SUBAPPLICATION Uebung_268_AX (* Race Condition mit E_SPLIT: zwei falsche und zwei richtige Varianten (Adapter) *)
  (* Standard: 61499-2; Description: Copyright (c) 2026 Meisterschulen am Ostbahnhof This program and the accompanying materials are made available under the terms of the Eclipse Public License 2.0 which is available at https://www.eclipse.org/legal/epl-2.0/ SPDX-License-Identifier: EPL-2.0 *)
  (* Version 1.0, 2026-11-11, Franz Höpfinger, Meisterschulen am Ostbahnhof, initial API and implementation and/or initial documentation *)
  PACKAGE Uebungen;
  IMPORT logiBUS::io::DI::logiBUS_DI::Input_I1;
  IMPORT logiBUS::io::DI::logiBUS_DI::Input_I2;
  IMPORT logiBUS::io::DI::logiBUS_DI::Input_I3;
  IMPORT logiBUS::io::DI::logiBUS_DI::Input_I4;
  IMPORT logiBUS::io::DI::logiBUS_DI_Events::BUTTON_SINGLE_CLICK;
  IMPORT logiBUS::io::DQ::logiBUS_DO::Output_Q1;
  IMPORT logiBUS::io::DQ::logiBUS_DO::Output_Q2;
  IMPORT logiBUS::io::DQ::logiBUS_DO::Output_Q3;
  IMPORT logiBUS::io::DQ::logiBUS_DO::Output_Q4;
  IMPORT logiBUS::io::DQ::logiBUS_DO::Output_Q5;
  IMPORT logiBUS::io::DQ::logiBUS_DO::Output_Q6;
  IMPORT logiBUS::io::DQ::logiBUS_DO::Output_Q7;
  IMPORT logiBUS::io::DQ::logiBUS_DO::Output_Q8;
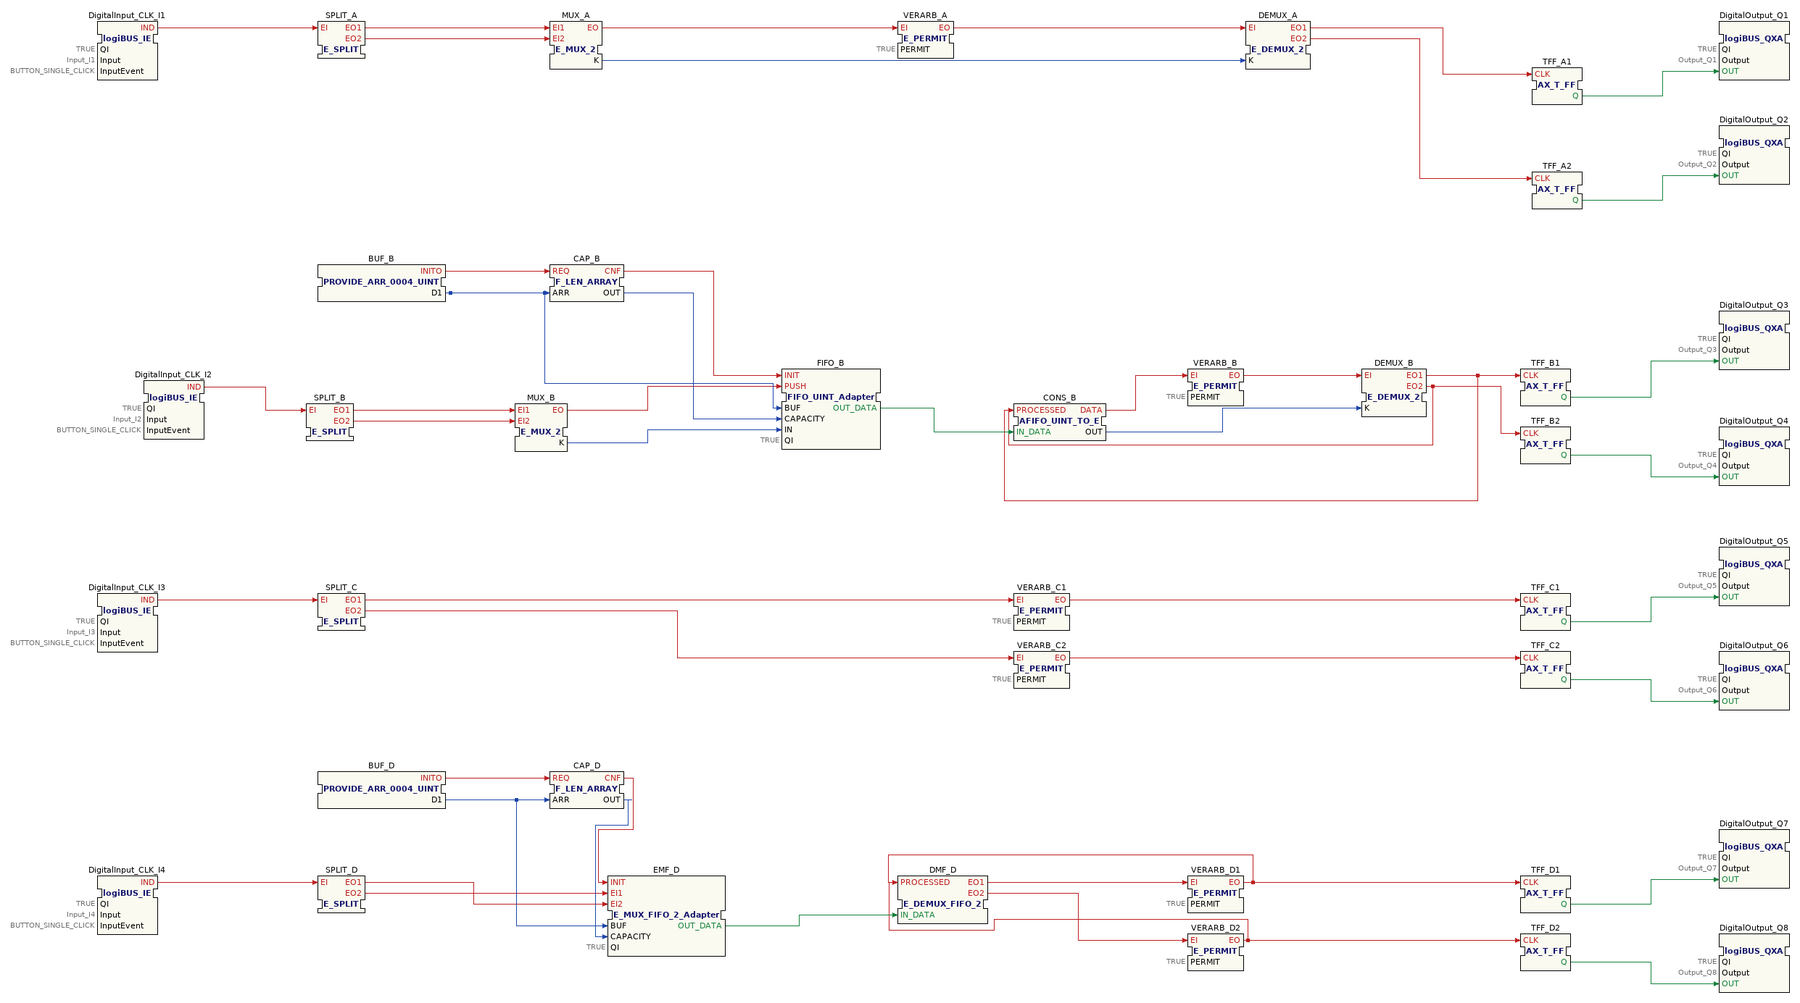
  FBS
    DigitalInput_CLK_I1 : logiBUS::io::DI::logiBUS_IE(QI := TRUE, Input := Input_I1, InputEvent := BUTTON_SINGLE_CLICK);
    SPLIT_A : iec61499::events::E_SPLIT;
    MUX_A : iec61499::events::E_MUX_2;
    VERARB_A : iec61499::events::E_PERMIT(PERMIT := TRUE);
    DEMUX_A : iec61499::events::E_DEMUX_2;
    TFF_A1 : adapter::events::unidirectional::AX_T_FF;
    DigitalOutput_Q1 : logiBUS::io::DQ::logiBUS_QXA(QI := TRUE, Output := Output_Q1);
    TFF_A2 : adapter::events::unidirectional::AX_T_FF;
    DigitalOutput_Q2 : logiBUS::io::DQ::logiBUS_QXA(QI := TRUE, Output := Output_Q2);
    DigitalInput_CLK_I2 : logiBUS::io::DI::logiBUS_IE(QI := TRUE, Input := Input_I2, InputEvent := BUTTON_SINGLE_CLICK);
    SPLIT_B : iec61499::events::E_SPLIT;
    BUF_B : eclipse4diac::convert::providers::PROVIDE_ARR_0004_UINT;
    CAP_B : eclipse4diac::utils::arrays::F_LEN_ARRAY;
    MUX_B : iec61499::events::E_MUX_2;
    FIFO_B : FIFO_adapter::FIFO_UINT_Adapter(QI := TRUE);
    CONS_B : FIFO_adapter::AFIFO_UINT_TO_E;
    VERARB_B : iec61499::events::E_PERMIT(PERMIT := TRUE);
    DEMUX_B : iec61499::events::E_DEMUX_2;
    TFF_B1 : adapter::events::unidirectional::AX_T_FF;
    DigitalOutput_Q3 : logiBUS::io::DQ::logiBUS_QXA(QI := TRUE, Output := Output_Q3);
    TFF_B2 : adapter::events::unidirectional::AX_T_FF;
    DigitalOutput_Q4 : logiBUS::io::DQ::logiBUS_QXA(QI := TRUE, Output := Output_Q4);
    DigitalInput_CLK_I3 : logiBUS::io::DI::logiBUS_IE(QI := TRUE, Input := Input_I3, InputEvent := BUTTON_SINGLE_CLICK);
    SPLIT_C : iec61499::events::E_SPLIT;
    VERARB_C1 : iec61499::events::E_PERMIT(PERMIT := TRUE);
    VERARB_C2 : iec61499::events::E_PERMIT(PERMIT := TRUE);
    TFF_C1 : adapter::events::unidirectional::AX_T_FF;
    DigitalOutput_Q5 : logiBUS::io::DQ::logiBUS_QXA(QI := TRUE, Output := Output_Q5);
    TFF_C2 : adapter::events::unidirectional::AX_T_FF;
    DigitalOutput_Q6 : logiBUS::io::DQ::logiBUS_QXA(QI := TRUE, Output := Output_Q6);
    DigitalInput_CLK_I4 : logiBUS::io::DI::logiBUS_IE(QI := TRUE, Input := Input_I4, InputEvent := BUTTON_SINGLE_CLICK);
    SPLIT_D : iec61499::events::E_SPLIT;
    BUF_D : eclipse4diac::convert::providers::PROVIDE_ARR_0004_UINT;
    CAP_D : eclipse4diac::utils::arrays::F_LEN_ARRAY;
    EMF_D : FIFO_adapter::E_MUX_FIFO_2_Adapter(QI := TRUE);
    DMF_D : FIFO_adapter::E_DEMUX_FIFO_2;
    VERARB_D1 : iec61499::events::E_PERMIT(PERMIT := TRUE);
    VERARB_D2 : iec61499::events::E_PERMIT(PERMIT := TRUE);
    TFF_D1 : adapter::events::unidirectional::AX_T_FF;
    DigitalOutput_Q7 : logiBUS::io::DQ::logiBUS_QXA(QI := TRUE, Output := Output_Q7);
    TFF_D2 : adapter::events::unidirectional::AX_T_FF;
    DigitalOutput_Q8 : logiBUS::io::DQ::logiBUS_QXA(QI := TRUE, Output := Output_Q8);
  END_FBS
  EVENT_CONNECTIONS
    DigitalInput_CLK_I1.IND TO SPLIT_A.EI;
    SPLIT_A.EO1 TO MUX_A.EI1;
    SPLIT_A.EO2 TO MUX_A.EI2;
    MUX_A.EO TO VERARB_A.EI;
    VERARB_A.EO TO DEMUX_A.EI;
    DEMUX_A.EO1 TO TFF_A1.CLK;
    DEMUX_A.EO2 TO TFF_A2.CLK;
    DigitalInput_CLK_I2.IND TO SPLIT_B.EI;
    BUF_B.INITO TO CAP_B.REQ;
    CAP_B.CNF TO FIFO_B.INIT;
    SPLIT_B.EO1 TO MUX_B.EI1;
    SPLIT_B.EO2 TO MUX_B.EI2;
    MUX_B.EO TO FIFO_B.PUSH;
    CONS_B.DATA TO VERARB_B.EI;
    VERARB_B.EO TO DEMUX_B.EI;
    DEMUX_B.EO1 TO CONS_B.PROCESSED;
    DEMUX_B.EO2 TO CONS_B.PROCESSED;
    DEMUX_B.EO1 TO TFF_B1.CLK;
    DEMUX_B.EO2 TO TFF_B2.CLK;
    DigitalInput_CLK_I3.IND TO SPLIT_C.EI;
    SPLIT_C.EO1 TO VERARB_C1.EI;
    SPLIT_C.EO2 TO VERARB_C2.EI;
    VERARB_C1.EO TO TFF_C1.CLK;
    VERARB_C2.EO TO TFF_C2.CLK;
    DigitalInput_CLK_I4.IND TO SPLIT_D.EI;
    BUF_D.INITO TO CAP_D.REQ;
    CAP_D.CNF TO EMF_D.INIT;
    SPLIT_D.EO1 TO EMF_D.EI1;
    SPLIT_D.EO2 TO EMF_D.EI2;
    DMF_D.EO1 TO VERARB_D1.EI;
    DMF_D.EO2 TO VERARB_D2.EI;
    VERARB_D1.EO TO DMF_D.PROCESSED;
    VERARB_D2.EO TO DMF_D.PROCESSED;
    VERARB_D1.EO TO TFF_D1.CLK;
    VERARB_D2.EO TO TFF_D2.CLK;
  END_CONNECTIONS
  DATA_CONNECTIONS
    MUX_A.K TO DEMUX_A.K;
    BUF_B.D1 TO CAP_B.ARR;
    BUF_B.D1 TO FIFO_B.BUF;
    CAP_B.OUT TO FIFO_B.CAPACITY;
    MUX_B.K TO FIFO_B.IN;
    CONS_B.OUT TO DEMUX_B.K;
    BUF_D.D1 TO CAP_D.ARR;
    BUF_D.D1 TO EMF_D.BUF;
    CAP_D.OUT TO EMF_D.CAPACITY;
  END_CONNECTIONS
  ADAPTER_CONNECTIONS
    TFF_A1.Q TO DigitalOutput_Q1.OUT;
    TFF_A2.Q TO DigitalOutput_Q2.OUT;
    FIFO_B.OUT_DATA TO CONS_B.IN_DATA;
    TFF_B1.Q TO DigitalOutput_Q3.OUT;
    TFF_B2.Q TO DigitalOutput_Q4.OUT;
    TFF_C1.Q TO DigitalOutput_Q5.OUT;
    TFF_C2.Q TO DigitalOutput_Q6.OUT;
    EMF_D.OUT_DATA TO DMF_D.IN_DATA;
    TFF_D1.Q TO DigitalOutput_Q7.OUT;
    TFF_D2.Q TO DigitalOutput_Q8.OUT;
  END_CONNECTIONS
END_SUBAPPLICATION
